(* IEC 61131-3 sources: llm-plc-st-eval/data/processed_v2_primera/gpt-4o/I3/zero_shot, 3 files *)

(* ---- ejec_1.st ---- *)
FUNCTION_BLOCK FB_Alarmas
VAR_INPUT
    alm1 : BOOL; // Alarma de prioridad alta
    alm2 : BOOL; // Alarma de prioridad media
    alm3 : BOOL; // Alarma de prioridad baja
    ack1 : BOOL; // Reconocimiento de alarma 1
    ack2 : BOOL; // Reconocimiento de alarma 2
    ack3 : BOOL; // Reconocimiento de alarma 3
END_VAR

VAR_OUTPUT
    sirena : BOOL; // Indica si la sirena está activa
    codigoAlm : INT; // Código de la alarma de mayor prioridad activa
END_VAR

VAR
    ret1 : BOOL; // Retención de la alarma 1
    ret2 : BOOL; // Retención de la alarma 2
    ret3 : BOOL; // Retención de la alarma 3
END_VAR

// Retención de alarmas
IF alm1 THEN
    ret1 := TRUE;
END_IF;

IF alm2 THEN
    ret2 := TRUE;
END_IF;

IF alm3 THEN
    ret3 := TRUE;
END_IF;

// Reconocimiento de alarmas
IF ack1 AND NOT alm1 THEN
    ret1 := FALSE;
END_IF;

IF ack2 AND NOT alm2 THEN
    ret2 := FALSE;
END_IF;

IF ack3 AND NOT alm3 THEN
    ret3 := FALSE;
END_IF;

// Determinación de la alarma de mayor prioridad
IF ret1 THEN
    codigoAlm := 1;
ELSIF ret2 THEN
    codigoAlm := 2;
ELSIF ret3 THEN
    codigoAlm := 3;
ELSE
    codigoAlm := 0;
END_IF;

// Activación de la sirena
sirena := ret1 OR ret2 OR ret3;

END_FUNCTION_BLOCK

(* ---- ejec_2.st ---- *)
FUNCTION_BLOCK FB_Alarmas
VAR_INPUT
    alm1 : BOOL; // Alarma de prioridad alta
    alm2 : BOOL; // Alarma de prioridad media
    alm3 : BOOL; // Alarma de prioridad baja
    ack1 : BOOL; // Reconocimiento de alarma 1
    ack2 : BOOL; // Reconocimiento de alarma 2
    ack3 : BOOL; // Reconocimiento de alarma 3
END_VAR

VAR_OUTPUT
    sirena : BOOL; // Indica si la sirena está activa
    codigoAlm : INT; // Código de la alarma de mayor prioridad activa
END_VAR

VAR
    retAlm1 : BOOL; // Retención de alarma 1
    retAlm2 : BOOL; // Retención de alarma 2
    retAlm3 : BOOL; // Retención de alarma 3
END_VAR

// Retención de alarmas
IF alm1 THEN
    retAlm1 := TRUE;
END_IF;

IF alm2 THEN
    retAlm2 := TRUE;
END_IF;

IF alm3 THEN
    retAlm3 := TRUE;
END_IF;

// Reconocimiento de alarmas
IF ack1 AND NOT alm1 THEN
    retAlm1 := FALSE;
END_IF;

IF ack2 AND NOT alm2 THEN
    retAlm2 := FALSE;
END_IF;

IF ack3 AND NOT alm3 THEN
    retAlm3 := FALSE;
END_IF;

// Determinación de la alarma de mayor prioridad
IF retAlm1 THEN
    codigoAlm := 1;
ELSIF retAlm2 THEN
    codigoAlm := 2;
ELSIF retAlm3 THEN
    codigoAlm := 3;
ELSE
    codigoAlm := 0;
END_IF;

// Activación de la sirena si hay alguna alarma retenida
sirena := retAlm1 OR retAlm2 OR retAlm3;

END_FUNCTION_BLOCK

(* ---- ejec_3.st ---- *)
FUNCTION_BLOCK FB_Alarmas
VAR_INPUT
    alm1 : BOOL; // Entrada de alarma de prioridad alta
    alm2 : BOOL; // Entrada de alarma de prioridad media
    alm3 : BOOL; // Entrada de alarma de prioridad baja
    ack1 : BOOL; // Reconocimiento de alarma 1
    ack2 : BOOL; // Reconocimiento de alarma 2
    ack3 : BOOL; // Reconocimiento de alarma 3
END_VAR

VAR_OUTPUT
    sirena : BOOL; // Salida para activar la sirena
    codigoAlm : INT; // Código de la alarma de mayor prioridad activa
END_VAR

VAR
    retAlm1 : BOOL; // Retención de alarma 1
    retAlm2 : BOOL; // Retención de alarma 2
    retAlm3 : BOOL; // Retención de alarma 3
END_VAR

// Retención de alarmas
IF alm1 THEN
    retAlm1 := TRUE;
END_IF;

IF alm2 THEN
    retAlm2 := TRUE;
END_IF;

IF alm3 THEN
    retAlm3 := TRUE;
END_IF;

// Reconocimiento de alarmas
IF ack1 AND NOT alm1 THEN
    retAlm1 := FALSE;
END_IF;

IF ack2 AND NOT alm2 THEN
    retAlm2 := FALSE;
END_IF;

IF ack3 AND NOT alm3 THEN
    retAlm3 := FALSE;
END_IF;

// Determinación del código de alarma de mayor prioridad
IF retAlm1 THEN
    codigoAlm := 1;
ELSIF retAlm2 THEN
    codigoAlm := 2;
ELSIF retAlm3 THEN
    codigoAlm := 3;
ELSE
    codigoAlm := 0;
END_IF;

// Activación de la sirena si hay alguna alarma retenida
sirena := retAlm1 OR retAlm2 OR retAlm3;

END_FUNCTION_BLOCK
